// GUI -> SPS mit Übernahme durch ParamApply.
{attribute 'pack_mode' := '1'}
TYPE ST_HmiParam :
STRUCT
    nPlanId : UDINT;
    stMaterial : ST_Material;
    fFeedOverride_pct : LREAL; // 0..100
    fSingleAxisVelo_pct : LREAL; // 0..100
END_STRUCT
END_TYPE

(* stored: Version 1.1.0.1
   DUT ST_HmiParam: Id {3b7040a0-38d0-4604-a124-e839b9cbfb00} *)
